{attribute 'qualified_only'}
{attribute 'strict'}
{attribute 'to_string'}
TYPE E_WordOrder :
(
    BigEndian       := 0,
    LittleEndian    := 1
) UINT;
END_TYPE

(* stored: Version 1.1.0.1
   DUT E_WordOrder: Id {f738e18a-49bb-4d42-a719-23c2f867c04d} *)
